(* PLC project TBEN_L5_PLC11.project, CODESYS CODESYS V3.5 SP21 Patch 1 *)
(* stored: creationDateTime 2026-11-07T15:35:07.3348543, modificationDateTime 2026-11-07T15:09:07.4034196 *)

// 1 index trong bảng dữ liệu giả lập của FB_MockRecordAccess
TYPE ST_MockParam :
STRUCT
    uiIndex : UINT;
    eAccess : E_IolAccess;
    uiLen   : UINT;                      // số byte của cả index
    abData  : ARRAY[0..63] OF BYTE;      // big-endian như trên dây
END_STRUCT
END_TYPE
